{attribute 'qualified_only'}
{attribute 'strict'}
{attribute 'to_string'}
TYPE eLightTemperature :
(
	WARM,
	NEUTRAL,
	COLD
);
END_TYPE

(* stored: Version 1.1.0.1
   DUT eLightTemperature: Id {5d20d888-4a19-456f-8a97-f7a4b57f15fc} *)
